Fanuc KAREL source: kb00134.KL

-- PROVISIONAL review KL for V770-1; original PC SHA256 cc89db503e2fe7bcea5151f60216f28e7cee5c4a50279e5622b9b8d0497c77e6
-- Incomplete behavior may be omitted. Consult companion uncertainty JSON. Do not deploy.
PROGRAM KB00134
%NOLOCKGROUP
BEGIN
  -- UNRESOLVED_PC offsets 5-12; opcodes 9D,23
  -- UNRESOLVED_PC offsets 17-26; opcodes 3F,75
  -- UNRESOLVED_PC offsets 31-38; opcodes 9D,23
  -- UNRESOLVED_PC offsets 43-50; opcodes 9D,23
  -- UNRESOLVED_PC offsets 55-85; opcodes 27,22,22,2A,22,22,31
  -- UNRESOLVED_PC offsets 90-94; opcodes 7F
END KB00134
